FUNCTION_BLOCK DlPgnRequest (* Send a request (PGN 59904) for a PGN *)
  (* Standard: 61499-2; Description: Calls iso_DlPgnRequest() of the CCI ISOBUS driver (data link layer, ISO 11783-3). \n No Rx PGN needs to be installed. The answer is received by an installed Rx PGN, if any. \n Sender is NmDestin.s16OwnCfHnd, receiver is NmDestin.s16Handle (HANDLE::GLOBAL for a global request). \n For PDU1 PGNs the lower byte of u32Pgn must be zero. *)
  (* Version 1.0, 2026-11-17, Franz Höpfinger, initial API and implementation and/or initial documentation *)
  PACKAGE isobus::pgn::tx;
  IMPORT isobus::pgn::ISONETEVENT_T;
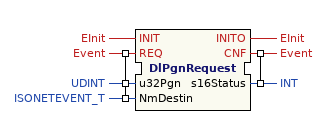
  EVENT_INPUT
    INIT : EInit; (* Service Initialization *)
    REQ WITH u32Pgn, NmDestin; (* Send the request *)
  END_EVENT
  EVENT_OUTPUT
    INITO : EInit; (* Initialization Confirm *)
    CNF WITH s16Status; (* Request sent (see s16Status) *)
  END_EVENT
  VAR_INPUT
    u32Pgn : UDINT; (* Requested PGN - Range: 0 - 0x3FFFF *)
    NmDestin : isobus::pgn::ISONETEVENT_T; (* Sender (s16OwnCfHnd) and receiver (s16Handle) *)
  END_VAR
  VAR_OUTPUT
    s16Status : INT; (* Return value of iso_DlPgnRequest(): 0 = OK *)
  END_VAR
END_FUNCTION_BLOCK
